(*
SPDX-FileCopyrightText: © 2026 Oleksandr Tiutyk <trofimich@gmail.com>
SPDX-License-Identifier: MIT
License: https://opensource.org/license/mit
*)

(*!
<summary>
Beckhoff incremental encoder input channel process image.
</summary>
<description>
Encapsulates 16-bit status word, 32-bit position value, and 32-bit captured latch value.
Use the matching 32-bit main PDO of EL5101 enhanced mode or EL5151. EL5152 has no latch and uses
INCREMENTAL_ENCODER_COUNTER_INPUT_CHANNEL instead; 16-bit process images are unsupported.
When used for I/O, link located fields or their containing buffers to the matching selected PDOs.
The record is not a packed wire buffer; compiler padding is not part of the device specification.
Unlinked/default values do not prove valid I/O. The caller evaluates bus/channel validity before use.
Use one owner task per instance and externally synchronize other access; multi-field snapshots are not atomic.
Copies store data without creating hardware links. Keep borrowed field references valid while consumers are bound.
This passive record performs no validation, synchronization, configuration or protocol advancement.
</description>
*)
TYPE INCREMENTAL_ENCODER_INPUT_CHANNEL :
STRUCT
	Status AT %I* : WORD;
	Value AT %I* : UDINT;
	Latch AT %I* : UDINT;
END_STRUCT
END_TYPE

(* stored: Version 1.1.0.1, ProductVersion 3.1.4026.20
   DUT INCREMENTAL_ENCODER_INPUT_CHANNEL: Id {6405443f-1275-4de4-a57c-09eb949b6716} *)
